(* IEC 61131-3 sources: llm-plc-st-eval/codesys/dobles/I7, 10 files *)

(* ---- 01_Correcta.st ---- *)
(* DOBLE DE PRUEBA I7/Correcta - NO ES CORPUS. Esperado: veredicto 1 *)
FUNCTION_BLOCK FB_Duplex
VAR_INPUT
    demanda : BOOL;
    falla1 : BOOL;
    falla2 : BOOL;
END_VAR
VAR_OUTPUT
    bomba1 : BOOL;
    bomba2 : BOOL;
    almFalla : BOOL;
END_VAR
VAR
    turno : BOOL;
    fDem : R_TRIG;
END_VAR
fDem(CLK := demanda);
IF fDem.Q THEN
    turno := NOT turno;
END_IF
IF demanda THEN
    IF turno THEN
        bomba1 := NOT falla1;
        bomba2 := falla1 AND NOT falla2;
        almFalla := falla1;
    ELSE
        bomba2 := NOT falla2;
        bomba1 := falla2 AND NOT falla1;
        almFalla := falla2;
    END_IF
ELSE
    bomba1 := FALSE;
    bomba2 := FALSE;
    almFalla := FALSE;
END_IF
END_FUNCTION_BLOCK

(* ---- 02_ReferenciaC4.st ---- *)
(* DOBLE DE PRUEBA I7/ReferenciaC4 - NO ES CORPUS. Esperado: veredicto 1 *)
FUNCTION_BLOCK FB_Duplex
VAR_INPUT
    demanda : BOOL;
    falla1 : BOOL;
    falla2 : BOOL;
END_VAR
VAR_OUTPUT
    bomba1 : BOOL;
    bomba2 : BOOL;
    almFalla : BOOL;
END_VAR
VAR
    turno : BOOL;
    fDem : R_TRIG;
END_VAR
fDem(CLK := demanda);
IF fDem.Q THEN
    turno := NOT turno;
END_IF
IF demanda THEN
    IF turno THEN
        bomba1 := NOT falla1;
        bomba2 := falla1 AND NOT falla2;
        almFalla := falla1;
    ELSE
        bomba2 := NOT falla2;
        bomba1 := falla2 AND NOT falla1;
        almFalla := falla2;
    END_IF
ELSE
    bomba1 := FALSE;
    bomba2 := FALSE;
    almFalla := FALSE;
END_IF
END_FUNCTION_BLOCK

(* ---- 03_SinAlternancia.st ---- *)
(* DOBLE DE PRUEBA I7/SinAlternancia - NO ES CORPUS. Esperado: veredicto 2, falla en el paso 3 *)
FUNCTION_BLOCK FB_Duplex
VAR_INPUT
    demanda : BOOL;
    falla1 : BOOL;
    falla2 : BOOL;
END_VAR
VAR_OUTPUT
    bomba1 : BOOL;
    bomba2 : BOOL;
    almFalla : BOOL;
END_VAR
VAR
    turno : BOOL;
    fDem : R_TRIG;
END_VAR
fDem(CLK := demanda);
turno := TRUE;
IF demanda THEN
    IF turno THEN
        bomba1 := NOT falla1;
        bomba2 := falla1 AND NOT falla2;
        almFalla := falla1;
    ELSE
        bomba2 := NOT falla2;
        bomba1 := falla2 AND NOT falla1;
        almFalla := falla2;
    END_IF
ELSE
    bomba1 := FALSE;
    bomba2 := FALSE;
    almFalla := FALSE;
END_IF
END_FUNCTION_BLOCK

(* ---- 04_PrimeraEsB2.st ---- *)
(* DOBLE DE PRUEBA I7/PrimeraEsB2 - NO ES CORPUS. Esperado: veredicto 2, falla en el paso 1 *)
FUNCTION_BLOCK FB_Duplex
VAR_INPUT
    demanda : BOOL;
    falla1 : BOOL;
    falla2 : BOOL;
END_VAR
VAR_OUTPUT
    bomba1 : BOOL;
    bomba2 : BOOL;
    almFalla : BOOL;
END_VAR
VAR
    turno : BOOL;
    fDem : R_TRIG;
END_VAR
fDem(CLK := demanda);
IF fDem.Q THEN
    turno := NOT turno;
END_IF
IF demanda THEN
    IF NOT turno THEN
        bomba1 := NOT falla1;
        bomba2 := falla1 AND NOT falla2;
        almFalla := falla1;
    ELSE
        bomba2 := NOT falla2;
        bomba1 := falla2 AND NOT falla1;
        almFalla := falla2;
    END_IF
ELSE
    bomba1 := FALSE;
    bomba2 := FALSE;
    almFalla := FALSE;
END_IF
END_FUNCTION_BLOCK

(* ---- 05_AmbasArrancan.st ---- *)
(* DOBLE DE PRUEBA I7/AmbasArrancan - NO ES CORPUS. Esperado: veredicto 2, falla en el paso 1 *)
FUNCTION_BLOCK FB_Duplex
VAR_INPUT
    demanda : BOOL;
    falla1 : BOOL;
    falla2 : BOOL;
END_VAR
VAR_OUTPUT
    bomba1 : BOOL;
    bomba2 : BOOL;
    almFalla : BOOL;
END_VAR
VAR
    turno : BOOL;
    fDem : R_TRIG;
END_VAR
fDem(CLK := demanda);
IF fDem.Q THEN
    turno := NOT turno;
END_IF
IF demanda THEN
    IF turno THEN
        bomba1 := NOT falla1;
        bomba2 := falla1 AND NOT falla2;
        almFalla := falla1;
    ELSE
        bomba2 := NOT falla2;
        bomba1 := falla2 AND NOT falla1;
        almFalla := falla2;
    END_IF
ELSE
    bomba1 := FALSE;
    bomba2 := FALSE;
    almFalla := FALSE;
END_IF
IF demanda THEN
    bomba1 := NOT falla1;
    bomba2 := NOT falla2;
END_IF
END_FUNCTION_BLOCK

(* ---- 06_SinRespaldo.st ---- *)
(* DOBLE DE PRUEBA I7/SinRespaldo - NO ES CORPUS. Esperado: veredicto 2, falla en el paso 6 *)
FUNCTION_BLOCK FB_Duplex
VAR_INPUT
    demanda : BOOL;
    falla1 : BOOL;
    falla2 : BOOL;
END_VAR
VAR_OUTPUT
    bomba1 : BOOL;
    bomba2 : BOOL;
    almFalla : BOOL;
END_VAR
VAR
    turno : BOOL;
    fDem : R_TRIG;
END_VAR
fDem(CLK := demanda);
IF fDem.Q THEN
    turno := NOT turno;
END_IF
IF demanda THEN
    IF turno THEN
        bomba1 := NOT falla1;
        bomba2 := falla1 AND NOT falla2;
        almFalla := falla1;
    ELSE
        bomba2 := NOT falla2;
        bomba1 := falla2 AND NOT falla1;
        almFalla := falla2;
    END_IF
ELSE
    bomba1 := FALSE;
    bomba2 := FALSE;
    almFalla := FALSE;
END_IF
IF turno THEN
    bomba2 := FALSE;
ELSE
    bomba1 := FALSE;
END_IF
END_FUNCTION_BLOCK

(* ---- 07_RespaldoEnclavado.st ---- *)
(* DOBLE DE PRUEBA I7/RespaldoEnclavado - NO ES CORPUS. Esperado: veredicto 2, falla en el paso 7 *)
FUNCTION_BLOCK FB_Duplex
VAR_INPUT
    demanda : BOOL;
    falla1 : BOOL;
    falla2 : BOOL;
END_VAR
VAR_OUTPUT
    bomba1 : BOOL;
    bomba2 : BOOL;
    almFalla : BOOL;
END_VAR
VAR
    turno : BOOL;
    fDem : R_TRIG;
    enResp : BOOL;
END_VAR
fDem(CLK := demanda);
IF fDem.Q THEN
    turno := NOT turno;
END_IF
IF NOT demanda THEN
    enResp := FALSE;
ELSIF (turno AND falla1) OR (NOT turno AND falla2) THEN
    enResp := TRUE;
END_IF
IF NOT demanda THEN
    bomba1 := FALSE;
    bomba2 := FALSE;
    almFalla := FALSE;
ELSIF enResp THEN
    IF turno THEN
        bomba1 := FALSE;
        bomba2 := NOT falla2;
        almFalla := falla1;
    ELSE
        bomba2 := FALSE;
        bomba1 := NOT falla1;
        almFalla := falla2;
    END_IF
ELSE
        IF turno THEN
            bomba1 := NOT falla1;
            bomba2 := falla1 AND NOT falla2;
            almFalla := falla1;
        ELSE
            bomba2 := NOT falla2;
            bomba1 := falla2 AND NOT falla1;
            almFalla := falla2;
        END_IF
END_IF
END_FUNCTION_BLOCK

(* ---- 08_AlarmaPorRespaldo.st ---- *)
(* DOBLE DE PRUEBA I7/AlarmaPorRespaldo - NO ES CORPUS. Esperado: veredicto 2, falla en el paso 8 *)
FUNCTION_BLOCK FB_Duplex
VAR_INPUT
    demanda : BOOL;
    falla1 : BOOL;
    falla2 : BOOL;
END_VAR
VAR_OUTPUT
    bomba1 : BOOL;
    bomba2 : BOOL;
    almFalla : BOOL;
END_VAR
VAR
    turno : BOOL;
    fDem : R_TRIG;
END_VAR
fDem(CLK := demanda);
IF fDem.Q THEN
    turno := NOT turno;
END_IF
IF demanda THEN
    IF turno THEN
        bomba1 := NOT falla1;
        bomba2 := falla1 AND NOT falla2;
        almFalla := falla1;
    ELSE
        bomba2 := NOT falla2;
        bomba1 := falla2 AND NOT falla1;
        almFalla := falla2;
    END_IF
ELSE
    bomba1 := FALSE;
    bomba2 := FALSE;
    almFalla := FALSE;
END_IF
almFalla := demanda AND (falla1 OR falla2);
END_FUNCTION_BLOCK

(* ---- 09_RespaldoConFalla.st ---- *)
(* DOBLE DE PRUEBA I7/RespaldoConFalla - NO ES CORPUS. Esperado: veredicto 2, falla en el paso 9 *)
FUNCTION_BLOCK FB_Duplex
VAR_INPUT
    demanda : BOOL;
    falla1 : BOOL;
    falla2 : BOOL;
END_VAR
VAR_OUTPUT
    bomba1 : BOOL;
    bomba2 : BOOL;
    almFalla : BOOL;
END_VAR
VAR
    turno : BOOL;
    fDem : R_TRIG;
END_VAR
fDem(CLK := demanda);
IF fDem.Q THEN
    turno := NOT turno;
END_IF
IF demanda THEN
    IF turno THEN
        bomba1 := NOT falla1;
        bomba2 := falla1 AND NOT falla2;
        almFalla := falla1;
    ELSE
        bomba2 := NOT falla2;
        bomba1 := falla2 AND NOT falla1;
        almFalla := falla2;
    END_IF
ELSE
    bomba1 := FALSE;
    bomba2 := FALSE;
    almFalla := FALSE;
END_IF
IF demanda THEN
    IF turno THEN
        bomba2 := falla1;
    ELSE
        bomba1 := falla2;
    END_IF
END_IF
END_FUNCTION_BLOCK

(* ---- 10_AlarmaSinDemanda.st ---- *)
(* DOBLE DE PRUEBA I7/AlarmaSinDemanda - NO ES CORPUS. Esperado: veredicto 2, falla en el paso 10 *)
FUNCTION_BLOCK FB_Duplex
VAR_INPUT
    demanda : BOOL;
    falla1 : BOOL;
    falla2 : BOOL;
END_VAR
VAR_OUTPUT
    bomba1 : BOOL;
    bomba2 : BOOL;
    almFalla : BOOL;
END_VAR
VAR
    turno : BOOL;
    fDem : R_TRIG;
END_VAR
fDem(CLK := demanda);
IF fDem.Q THEN
    turno := NOT turno;
END_IF
IF demanda THEN
    IF turno THEN
        bomba1 := NOT falla1;
        bomba2 := falla1 AND NOT falla2;
        almFalla := falla1;
    ELSE
        bomba2 := NOT falla2;
        bomba1 := falla2 AND NOT falla1;
        almFalla := falla2;
    END_IF
ELSE
    bomba1 := FALSE;
    bomba2 := FALSE;
    almFalla := FALSE;
END_IF
IF turno THEN
    almFalla := falla1;
ELSE
    almFalla := falla2;
END_IF
END_FUNCTION_BLOCK
